(* IEC 61131-3 sources: SRCI_CLIENT_PLC/RobotLibrary/Library/POUs/Additional/MC_PathAccuracyMode/Structures, 4 files *)

(* ---- PathAccuracyModeOutCmd.st ---- *)
{attribute 'pack_mode' := '1'}
// -------------------------------------------------------------------------
//  SRCI Robot Library
// -------------------------------------------------------------------------
//
//  Object:      PathAccuracyModeOutCmd
//  Author:      Thorsten Brach
//  Date:        2024-06-22
//
//  Description:
//
//
//  Copyright:
//    (C) 2024 Thorsten Brach. All rights reserved
//             Licensed under the MIT License.
//
//  Disclaimer:
//    This project is provided without any guarantee and can be used for
//    private and commercial purposes. Any use is at the user’s
//    own risk and responsibility.
//
// -------------------------------------------------------------------------
TYPE PathAccuracyModeOutCmd :
STRUCT
END_STRUCT
END_TYPE

(* ---- PathAccuracyModeParCmd.st ---- *)
{attribute 'pack_mode' := '1'}
// -------------------------------------------------------------------------
//  SRCI Robot Library
// -------------------------------------------------------------------------
//
//  Object:      PathAccuracyModeParCmd
//  Author:      Thorsten Brach
//  Date:        2024-06-22
//
//  Description:
//
//
//  Copyright:
//    (C) 2024 Thorsten Brach. All rights reserved
//             Licensed under the MIT License.
//
//  Disclaimer:
//    This project is provided without any guarantee and can be used for
//    private and commercial purposes. Any use is at the user’s
//    own risk and responsibility.
//
// -------------------------------------------------------------------------
TYPE PathAccuracyModeParCmd :
STRUCT
END_STRUCT
END_TYPE

(* ---- PathAccuracyModeRecvData.st ---- *)
{attribute 'pack_mode' := '1'}
// -------------------------------------------------------------------------
//  SRCI Robot Library
// -------------------------------------------------------------------------
//
//  Object:      PathAccuracyModeRecvData
//  Author:      Thorsten Brach
//  Date:        2024-06-22
//
//  Description:
//
//
//  Copyright:
//    (C) 2024 Thorsten Brach. All rights reserved
//             Licensed under the MIT License.
//
//  Disclaimer:
//    This project is provided without any guarantee and can be used for
//    private and commercial purposes. Any use is at the user’s
//    own risk and responsibility.
//
// -------------------------------------------------------------------------
TYPE PathAccuracyModeRecvData EXTENDS RspHeader :
STRUCT
  /// TRUE while PathAccuracyMode is active
  Enabled : BOOL;
END_STRUCT
END_TYPE

(* ---- PathAccuracyModeSendData.st ---- *)
{attribute 'pack_mode' := '1'}
// -------------------------------------------------------------------------
//  SRCI Robot Library
// -------------------------------------------------------------------------
//
//  Object:      PathAccuracyModeSendData
//  Author:      Thorsten Brach
//  Date:        2024-06-22
//
//  Description:
//
//
//  Copyright:
//    (C) 2024 Thorsten Brach. All rights reserved
//             Licensed under the MIT License.
//
//  Disclaimer:
//    This project is provided without any guarantee and can be used for
//    private and commercial purposes. Any use is at the user’s
//    own risk and responsibility.
//
// -------------------------------------------------------------------------
TYPE PathAccuracyModeSendData EXTENDS CmdHeader:
STRUCT
  /// Set TRUE to activate monitoring of work areas
  Enable             : BOOL;
END_STRUCT
END_TYPE
